(* IEC 61131-3 sources: s7-to-codesys/s7conv/tests/snapshots/fixtures/src/GVLs, 6 files *)

(* ---- DB_Hmi.gvl.st ---- *)
// Назначение: Глобальный DB «DB_Hmi», сконвертирован из SCL
// Автор:      не указан (исходный блок S7); перевод в ST — s7conv 0.1.0
// Версия:     0.1 (исходный блок S7)
// Документ:   docs/CONVERSION_REPORT.md, docs/MAPPING.md
// Источник:   s7conv/tests/fixtures/main.scl, строки 43–54, DATA_BLOCK "DB_Hmi"
// Сгенерировано s7conv: пометки MIGRATION-CHECK и MIGRATION-TODO требуют ручного разбора.
{attribute 'qualified_only'}
VAR_GLOBAL
    ackRequest : BOOL;
    counter : INT;
END_VAR

(* ---- DB_Settings.gvl.st ---- *)
// Назначение: Глобальный DB «DB_Settings», сконвертирован из SCL
// Автор:      не указан (исходный блок S7); перевод в ST — s7conv 0.1.0
// Версия:     0.1 (исходный блок S7)
// Документ:   docs/CONVERSION_REPORT.md, docs/MAPPING.md
// Источник:   s7conv/tests/fixtures/analog.scl, строки 31–48, DATA_BLOCK "DB_Settings"
// Сгенерировано s7conv: пометки MIGRATION-CHECK и MIGRATION-TODO требуют ручного разбора.
{attribute 'qualified_only'}
VAR_GLOBAL
    levelLow : REAL := 0.0;
    levelHigh : REAL := 95.5;
    pumpDelay : TIME := T#5s;
    // MIGRATION-CHECK: S5Time → TIME: в S7 S5TIME — BCD с шагом 10 мс…10 с, диапазон до 2h46m30s (стр. 38)
    oldDelay : TIME := T#2s;
    label : STRING(254);
END_VAR
VAR_GLOBAL RETAIN
    totalVolume : LREAL;
    counterRaw : INT;
END_VAR

(* ---- GVL_InstanceDBs.gvl.st ---- *)
// Назначение: экземпляры функциональных блоков и типизированные DB S7 (экземплярные DB → переменные GVL)
// Автор:      s7conv 0.1.0 (сгенерировано)
// Версия:     не указана
// Документ:   docs/MAPPING.md, раздел «DB»
{attribute 'qualified_only'}
VAR_GLOBAL
    Delay_DB : TON; // s7conv/tests/fixtures/main.scl:56
    Level_DB : FB_Level; // s7conv/tests/fixtures/main.scl:66
    Motor1_DB : FB_Motor; // s7conv/tests/fixtures/motor.scl:103
    // MIGRATION-CHECK: экземплярный DB FB_Legacy_DB выведен по вызову (исходника DB в корпусе нет)
    FB_Legacy_DB : FB_Legacy;
END_VAR

(* ---- GVL_IO.gvl.st ---- *)
// Назначение: символьный слой входов/выходов S7: прямые адреса и теги с адресом → переменные с AT
// Автор:      s7conv 0.1.0 (сгенерировано)
// Версия:     не указана
// Документ:   docs/MAPPING.md, раздел «Адреса»
// Адресная модель: S7 нумерует байты (%IW64 — байты 64–65, big-endian), CODESYS — слова
// (%IW32 — байты 64–65, little-endian). Адреса ниже — заготовка: на ПЛК210 каналы модулей
// привязываются в дереве устройств (I/O mapping) — сверить с конфигурацией.
{attribute 'qualified_only'}
VAR_GLOBAL
    Start_PB AT %IX0.0 : BOOL; // S7 %I0.0; Кнопка «Пуск»
    Stop_PB AT %IX0.1 : BOOL; // S7 %I0.1; Кнопка «Стоп» (NC)
    I0_2 AT %IX0.2 : BOOL; // S7 %I0.2
    Level_Raw AT %IW32 : INT; // S7 %IW64; Уровень, сырое значение
    Motor_Run AT %QX0.0 : BOOL; // S7 %Q0.0; Пускатель двигателя
    Horn AT %QX0.1 : BOOL; // S7 %Q0.1; Сирена
    Q4_0 AT %QX4.0 : BOOL; // S7 %Q4.0
END_VAR

(* ---- GVL_Markers.gvl.st ---- *)
// Назначение: символьный слой меркеров (%M) S7: прямые адреса и теги с адресом → переменные с AT
// Автор:      s7conv 0.1.0 (сгенерировано)
// Версия:     не указана
// Документ:   docs/MAPPING.md, раздел «Адреса»
// Адресная модель: S7 нумерует байты (%IW64 — байты 64–65, big-endian), CODESYS — слова
// (%IW32 — байты 64–65, little-endian). Адреса ниже — заготовка: на ПЛК210 каналы модулей
// привязываются в дереве устройств (I/O mapping) — сверить с конфигурацией.
{attribute 'qualified_only'}
VAR_GLOBAL
    MW10 AT %MW5 : WORD; // S7 %MW10
    M12_1 AT %MX12.1 : BOOL; // S7 %M12.1
END_VAR

(* ---- GVL_Tags.gvl.st ---- *)
// Назначение: глобальные теги S7 без адреса и символы, не найденные в корпусе
// Автор:      s7conv 0.1.0 (сгенерировано)
// Версия:     не указана
// Документ:   docs/MAPPING.md, раздел «Теги»
{attribute 'qualified_only'}
VAR_GLOBAL
    // MIGRATION-CHECK: символ "Alarm_Lamp" не найден — тип BOOL выведен по использованию
    //                  (s7conv/tests/fixtures/analog.scl:69)
    Alarm_Lamp : BOOL;
END_VAR
